(* IEC 61131-3 sources: plcc/demo/st-programs, 7 files *)

(* ---- alarm_system.st ---- *)
FUNCTION PriorityEncode : INT
VAR_INPUT critical : INT; high : INT; medium : INT; low : INT; END_VAR
    IF critical <> 0 THEN PriorityEncode := 4;
    ELSIF high <> 0 THEN PriorityEncode := 3;
    ELSIF medium <> 0 THEN PriorityEncode := 2;
    ELSIF low <> 0 THEN PriorityEncode := 1;
    ELSE PriorityEncode := 0;
    END_IF;
END_FUNCTION

FUNCTION_BLOCK AlarmHandler
VAR_INPUT
    temp_alarm : BOOL;
    pressure_alarm : BOOL;
    level_alarm : BOOL;
END_VAR
VAR_OUTPUT
    alarm_active : BOOL;
    alarm_code : INT;
END_VAR
VAR
    temp_val : INT;
    press_val : INT;
    level_val : INT;
END_VAR
    IF temp_alarm THEN temp_val := 1; ELSE temp_val := 0; END_IF;
    IF pressure_alarm THEN press_val := 1; ELSE press_val := 0; END_IF;
    IF level_alarm THEN level_val := 1; ELSE level_val := 0; END_IF;
    alarm_code := PriorityEncode(press_val, temp_val, level_val, 0);
    alarm_active := alarm_code > 0;
END_FUNCTION_BLOCK

PROGRAM AlarmSystem
VAR
    handler : AlarmHandler;
    system_alarm : BOOL;
    system_code : INT;
END_VAR
    handler(temp_alarm := TRUE, pressure_alarm := FALSE, level_alarm := TRUE);
    system_alarm := handler.alarm_active;
    system_code := handler.alarm_code;
END_PROGRAM

(* ---- motor_control.st ---- *)
FUNCTION_BLOCK MotorController
VAR_INPUT
    start_cmd : BOOL;
    stop_cmd : BOOL;
    current : REAL;
    overload_limit : REAL := 15.0;
END_VAR
VAR_OUTPUT
    running : BOOL;
    fault : BOOL;
    run_time : INT;
END_VAR
VAR
    overload_count : INT := 0;
END_VAR
    IF stop_cmd OR fault THEN
        running := FALSE;
    ELSIF start_cmd AND NOT fault THEN
        running := TRUE;
    END_IF;

    IF running THEN
        run_time := run_time + 1;
        IF current > overload_limit THEN
            overload_count := overload_count + 1;
            IF overload_count >= 3 THEN
                fault := TRUE;
                running := FALSE;
            END_IF;
        ELSE
            overload_count := 0;
        END_IF;
    END_IF;
END_FUNCTION_BLOCK

PROGRAM MotorSystem
VAR
    motor1 : MotorController;
    motor2 : MotorController;
    any_fault : BOOL;
END_VAR
    motor1(start_cmd := TRUE, stop_cmd := FALSE, current := 10.0);
    motor2(start_cmd := TRUE, stop_cmd := FALSE, current := 10.0);
    any_fault := motor1.fault OR motor2.fault;
END_PROGRAM

(* ---- pid_simple.st ---- *)
FUNCTION_BLOCK PID
VAR_INPUT
    setpoint : REAL;
    measured : REAL;
    kp : REAL := 1.0;
    ki : REAL := 0.1;
    kd : REAL := 0.05;
    dt : REAL := 0.01;
    out_min : REAL := -100.0;
    out_max : REAL := 100.0;
END_VAR
VAR_OUTPUT
    output : REAL;
END_VAR
VAR
    err : REAL;
    prev_err : REAL := 0.0;
    integral : REAL := 0.0;
    derivative : REAL;
END_VAR
    err := setpoint - measured;
    integral := integral + err * dt;
    derivative := (err - prev_err) / dt;
    output := kp * err + ki * integral + kd * derivative;

    (* Clamp output *)
    IF output > out_max THEN
        output := out_max;
    ELSIF output < out_min THEN
        output := out_min;
    END_IF;

    prev_err := err;
END_FUNCTION_BLOCK

PROGRAM PIDController
VAR
    pid_inst : PID;
    sensor_value : REAL := 0.0;
    target_value : REAL := 50.0;
    control_output : REAL;
END_VAR
    pid_inst(setpoint := target_value, measured := sensor_value);
    control_output := pid_inst.output;
END_PROGRAM

(* ---- water_treatment.st ---- *)
(* ═══════════════════════════════════════════════════════════ *)
(*  Water Treatment Plant — Industrial PLC Program            *)
(*  Registers 0-39 are SCADA-accessible via Modbus            *)
(* ═══════════════════════════════════════════════════════════ *)

(* ── Function Blocks ── *)

FUNCTION_BLOCK TankLevel
VAR_INPUT
    inlet_flow : REAL;
    outlet_flow : REAL;
    max_capacity : REAL;
END_VAR
VAR_OUTPUT
    level : REAL;
    level_pct : INT;
    high_alarm : BOOL;
    low_alarm : BOOL;
END_VAR
VAR
    high_sp : REAL := 90.0;
    low_sp : REAL := 10.0;
END_VAR
    level := level + (inlet_flow - outlet_flow) * 0.001;
    IF level < 0.0 THEN level := 0.0; END_IF;
    IF level > max_capacity THEN level := max_capacity; END_IF;
    level_pct := REAL_TO_INT(level * 100.0 / max_capacity);
    high_alarm := level_pct > 90;
    low_alarm := level_pct < 10;
END_FUNCTION_BLOCK

FUNCTION_BLOCK PumpControl
VAR_INPUT
    cmd_start : BOOL;
    cmd_stop : BOOL;
    speed_sp : INT;
    fault_reset : BOOL;
END_VAR
VAR_OUTPUT
    running : BOOL;
    speed : INT;
    fault : BOOL;
    hours : INT;
END_VAR
VAR
    scans : INT := 0;
END_VAR
    IF fault_reset THEN fault := FALSE; END_IF;
    IF cmd_stop THEN running := FALSE; END_IF;
    IF cmd_start AND NOT fault THEN running := TRUE; END_IF;
    IF running THEN
        speed := speed_sp;
        scans := scans + 1;
        hours := scans / 3600;
    ELSE
        speed := 0;
    END_IF;
END_FUNCTION_BLOCK

FUNCTION_BLOCK ValveControl
VAR_INPUT
    cmd_open : BOOL;
    cmd_close : BOOL;
END_VAR
VAR_OUTPUT
    position : INT;
    opened : BOOL;
    closed : BOOL;
END_VAR
    IF cmd_open AND NOT cmd_close THEN
        IF position < 100 THEN position := position + 5; END_IF;
    ELSIF cmd_close AND NOT cmd_open THEN
        IF position > 0 THEN position := position - 5; END_IF;
    END_IF;
    opened := position >= 100;
    closed := position <= 0;
END_FUNCTION_BLOCK

(* ── Main Program ── *)

PROGRAM WaterTreatment
VAR
    (* ═══════════════════════════════════════════ *)
    (* COMMANDS — write from SCADA (R0-R9)        *)
    (* ═══════════════════════════════════════════ *)
    cmd_start : INT := 0;         (* R0  write 1 to start *)
    cmd_stop : INT := 0;          (* R1  write 1 to stop *)
    cmd_flush : INT := 0;         (* R2  write 1 to flush *)
    cmd_alarm_ack : INT := 0;     (* R3  write 1 to acknowledge alarms *)
    cmd_alarm_reset : INT := 0;   (* R4  write 1 to reset faults *)
    sp_raw_tank : INT := 50;      (* R5  raw tank level setpoint % *)
    sp_clean_tank : INT := 70;    (* R6  clean tank level setpoint % *)
    sp_inlet_pump : INT := 60;    (* R7  inlet pump speed % *)
    sp_transfer_pump : INT := 40; (* R8  transfer pump speed % *)
    sp_outlet_pump : INT := 30;   (* R9  outlet pump speed % *)

    (* ═══════════════════════════════════════════ *)
    (* STATUS — read from SCADA (R10-R19)         *)
    (* ═══════════════════════════════════════════ *)
    running : INT := 0;           (* R10 process running *)
    stopped : INT := 1;           (* R11 process stopped *)
    flushing : INT := 0;          (* R12 flush in progress *)
    faulted : INT := 0;           (* R13 fault/alarm state *)
    cycle_count : INT := 0;       (* R14 scan counter *)
    raw_level : INT := 0;         (* R15 raw tank level % *)
    clean_level : INT := 0;       (* R16 clean tank level % *)
    system_ok : INT := 1;         (* R17 all systems healthy *)
    alarm_word : INT := 0;        (* R18 alarm bitmask *)
    total_flow : INT := 0;        (* R19 cumulative output *)

    (* ═══════════════════════════════════════════ *)
    (* EQUIPMENT STATUS (R20-R31)                 *)
    (* ═══════════════════════════════════════════ *)
    inlet_pump_run : INT := 0;    (* R20 *)
    inlet_pump_speed : INT := 0;  (* R21 *)
    inlet_pump_fault : INT := 0;  (* R22 *)
    xfer_pump_run : INT := 0;     (* R23 *)
    xfer_pump_speed : INT := 0;   (* R24 *)
    xfer_pump_fault : INT := 0;   (* R25 *)
    outlet_pump_run : INT := 0;   (* R26 *)
    outlet_pump_speed : INT := 0; (* R27 *)
    outlet_pump_fault : INT := 0; (* R28 *)
    inlet_vlv_pos : INT := 0;     (* R29 *)
    outlet_vlv_pos : INT := 0;    (* R30 *)
    drain_vlv_pos : INT := 0;     (* R31 *)

    (* ═══════════════════════════════════════════ *)
    (* ALARMS (R32-R39)                           *)
    (* ═══════════════════════════════════════════ *)
    alm_raw_high : INT := 0;      (* R32 raw tank high level *)
    alm_raw_low : INT := 0;       (* R33 raw tank low level *)
    alm_clean_high : INT := 0;    (* R34 clean tank high level *)
    alm_clean_low : INT := 0;     (* R35 clean tank low level *)
    alm_inlet_fault : INT := 0;   (* R36 inlet pump fault *)
    alm_xfer_fault : INT := 0;    (* R37 transfer pump fault *)
    alm_outlet_fault : INT := 0;  (* R38 outlet pump fault *)
    alm_count : INT := 0;         (* R39 total active alarms *)

    (* ═══════════════════════════════════════════ *)
    (* INTERNAL — FB instances after registers     *)
    (* ═══════════════════════════════════════════ *)
    raw_tank : TankLevel;
    clean_tank : TankLevel;
    p_inlet : PumpControl;
    p_transfer : PumpControl;
    p_outlet : PumpControl;
    v_inlet : ValveControl;
    v_outlet : ValveControl;
    v_drain : ValveControl;

    prev_running : INT := -1;
    init_done : INT := 0;
END_VAR

    (* ── Startup ── *)
    IF init_done = 0 THEN
        PRINT('Water Treatment PLC started');
        init_done := 1;
    END_IF;
    cycle_count := cycle_count + 1;

    (* ── Process commands (edge-triggered, auto-clear) ── *)
    IF cmd_start = 1 THEN
        cmd_start := 0;
        IF faulted = 0 THEN
            running := 1; stopped := 0; flushing := 0;
            PRINT('CMD: Process START');
        END_IF;
    END_IF;

    IF cmd_stop = 1 THEN
        cmd_stop := 0;
        running := 0; stopped := 1; flushing := 0;
        PRINT('CMD: Process STOP');
    END_IF;

    IF cmd_flush = 1 THEN
        cmd_flush := 0;
        running := 0; stopped := 0; flushing := 1;
        PRINT('CMD: FLUSH started');
    END_IF;

    IF cmd_alarm_ack = 1 THEN
        cmd_alarm_ack := 0;
        PRINT('CMD: Alarms acknowledged');
    END_IF;

    IF cmd_alarm_reset = 1 THEN
        cmd_alarm_reset := 0;
        faulted := 0;
        system_ok := 1;
        p_inlet(cmd_start := FALSE, cmd_stop := FALSE, speed_sp := 0, fault_reset := TRUE);
        p_transfer(cmd_start := FALSE, cmd_stop := FALSE, speed_sp := 0, fault_reset := TRUE);
        p_outlet(cmd_start := FALSE, cmd_stop := FALSE, speed_sp := 0, fault_reset := TRUE);
        PRINT('CMD: Faults reset');
    END_IF;

    (* ── Process control ── *)
    IF running = 1 THEN
        (* Inlet: fill raw tank to setpoint *)
        IF raw_level < sp_raw_tank THEN
            p_inlet(cmd_start := TRUE, cmd_stop := FALSE, speed_sp := sp_inlet_pump, fault_reset := FALSE);
            v_inlet(cmd_open := TRUE, cmd_close := FALSE);
        ELSE
            p_inlet(cmd_start := FALSE, cmd_stop := TRUE, speed_sp := 0, fault_reset := FALSE);
            v_inlet(cmd_open := FALSE, cmd_close := TRUE);
        END_IF;

        (* Transfer: move water from raw to clean *)
        IF raw_level > 20 AND clean_level < sp_clean_tank THEN
            p_transfer(cmd_start := TRUE, cmd_stop := FALSE, speed_sp := sp_transfer_pump, fault_reset := FALSE);
        ELSE
            p_transfer(cmd_start := FALSE, cmd_stop := TRUE, speed_sp := 0, fault_reset := FALSE);
        END_IF;

        (* Outlet: distribute clean water *)
        IF clean_level > 30 THEN
            p_outlet(cmd_start := TRUE, cmd_stop := FALSE, speed_sp := sp_outlet_pump, fault_reset := FALSE);
            v_outlet(cmd_open := TRUE, cmd_close := FALSE);
        ELSE
            p_outlet(cmd_start := FALSE, cmd_stop := TRUE, speed_sp := 0, fault_reset := FALSE);
            v_outlet(cmd_open := FALSE, cmd_close := TRUE);
        END_IF;

        v_drain(cmd_open := FALSE, cmd_close := TRUE);

    ELSIF flushing = 1 THEN
        (* Flush: drain everything *)
        p_inlet(cmd_start := FALSE, cmd_stop := TRUE, speed_sp := 0, fault_reset := FALSE);
        p_transfer(cmd_start := FALSE, cmd_stop := TRUE, speed_sp := 0, fault_reset := FALSE);
        p_outlet(cmd_start := FALSE, cmd_stop := TRUE, speed_sp := 0, fault_reset := FALSE);
        v_inlet(cmd_open := FALSE, cmd_close := TRUE);
        v_outlet(cmd_open := FALSE, cmd_close := TRUE);
        v_drain(cmd_open := TRUE, cmd_close := FALSE);

        (* Auto-stop flush when tanks are empty *)
        IF raw_level = 0 AND clean_level = 0 THEN
            flushing := 0; stopped := 1;
            PRINT('Flush complete');
        END_IF;

    ELSE
        (* Stopped / faulted *)
        p_inlet(cmd_start := FALSE, cmd_stop := TRUE, speed_sp := 0, fault_reset := FALSE);
        p_transfer(cmd_start := FALSE, cmd_stop := TRUE, speed_sp := 0, fault_reset := FALSE);
        p_outlet(cmd_start := FALSE, cmd_stop := TRUE, speed_sp := 0, fault_reset := FALSE);
        v_inlet(cmd_open := FALSE, cmd_close := TRUE);
        v_outlet(cmd_open := FALSE, cmd_close := TRUE);
        v_drain(cmd_open := FALSE, cmd_close := TRUE);
    END_IF;

    (* ── Tank simulation ── *)
    (* Flow rates scaled for demo speed — tanks fill in ~30 seconds *)
    raw_tank(
        inlet_flow := INT_TO_REAL(p_inlet.speed) * 50.0,
        outlet_flow := INT_TO_REAL(p_transfer.speed) * 30.0,
        max_capacity := 1000.0
    );
    clean_tank(
        inlet_flow := INT_TO_REAL(p_transfer.speed) * 30.0,
        outlet_flow := INT_TO_REAL(p_outlet.speed) * 20.0,
        max_capacity := 500.0
    );

    (* ── Copy to SCADA registers ── *)
    raw_level := raw_tank.level_pct;
    clean_level := clean_tank.level_pct;

    inlet_pump_run := BOOL_TO_INT(p_inlet.running);
    inlet_pump_speed := p_inlet.speed;
    inlet_pump_fault := BOOL_TO_INT(p_inlet.fault);

    xfer_pump_run := BOOL_TO_INT(p_transfer.running);
    xfer_pump_speed := p_transfer.speed;
    xfer_pump_fault := BOOL_TO_INT(p_transfer.fault);

    outlet_pump_run := BOOL_TO_INT(p_outlet.running);
    outlet_pump_speed := p_outlet.speed;
    outlet_pump_fault := BOOL_TO_INT(p_outlet.fault);

    inlet_vlv_pos := v_inlet.position;
    outlet_vlv_pos := v_outlet.position;
    drain_vlv_pos := v_drain.position;

    total_flow := total_flow + p_outlet.speed;

    (* ── Alarms ── *)
    alm_raw_high := BOOL_TO_INT(raw_tank.high_alarm);
    alm_raw_low := BOOL_TO_INT(raw_tank.low_alarm);
    alm_clean_high := BOOL_TO_INT(clean_tank.high_alarm);
    alm_clean_low := BOOL_TO_INT(clean_tank.low_alarm);
    alm_inlet_fault := BOOL_TO_INT(p_inlet.fault);
    alm_xfer_fault := BOOL_TO_INT(p_transfer.fault);
    alm_outlet_fault := BOOL_TO_INT(p_outlet.fault);

    (* Alarm word: bitmask of all active alarms *)
    alarm_word := alm_raw_high + alm_raw_low * 2 + alm_clean_high * 4
                + alm_clean_low * 8 + alm_inlet_fault * 16
                + alm_xfer_fault * 32 + alm_outlet_fault * 64;

    alm_count := alm_raw_high + alm_raw_low + alm_clean_high + alm_clean_low
               + alm_inlet_fault + alm_xfer_fault + alm_outlet_fault;

    (* Trip to fault only on critical alarms: high level or pump faults *)
    (* Low level alarms are informational — not a fault condition *)
    IF running = 1 THEN
        IF alm_raw_high = 1 OR alm_clean_high = 1 OR alm_inlet_fault = 1 OR alm_xfer_fault = 1 OR alm_outlet_fault = 1 THEN
            faulted := 1;
            running := 0;
            system_ok := 0;
            PRINT('FAULT: critical alarm, process stopped');
        END_IF;
    END_IF;

END_PROGRAM

(* ---- batch_process.st ---- *)
PROGRAM BatchProcess
VAR
    stage : INT := 0;
    timer : INT := 0;
    fill_valve : BOOL := FALSE;
    mixer : BOOL := FALSE;
    drain_valve : BOOL := FALSE;
    batch_count : INT := 0;
    complete : BOOL := FALSE;
END_VAR
    timer := timer + 1;
    CASE stage OF
        0: (* IDLE *)
            fill_valve := FALSE; mixer := FALSE; drain_valve := FALSE;
            stage := 1; timer := 0;
        1: (* FILL *)
            fill_valve := TRUE;
            IF timer >= 20 THEN stage := 2; timer := 0; fill_valve := FALSE; END_IF;
        2: (* MIX *)
            mixer := TRUE;
            IF timer >= 30 THEN stage := 3; timer := 0; mixer := FALSE; END_IF;
        3: (* DRAIN *)
            drain_valve := TRUE;
            IF timer >= 15 THEN
                stage := 0; timer := 0; drain_valve := FALSE;
                batch_count := batch_count + 1;
                complete := TRUE;
            END_IF;
    ELSE
        stage := 0;
    END_CASE;
END_PROGRAM

(* ---- blink.st ---- *)
PROGRAM Blink
VAR
    output : BOOL := FALSE;
END_VAR
    output := NOT output;
END_PROGRAM

(* ---- state_machine.st ---- *)
PROGRAM StateMachine
VAR
    state : INT := 0;
    output_a : BOOL := FALSE;
    output_b : BOOL := FALSE;
    input_trigger : BOOL := FALSE;
    counter : INT := 0;
END_VAR
    CASE state OF
        0:
            output_a := FALSE;
            output_b := FALSE;
            IF input_trigger THEN
                state := 1;
            END_IF;
        1:
            output_a := TRUE;
            output_b := FALSE;
            counter := counter + 1;
            IF counter >= 10 THEN
                state := 2;
                counter := 0;
            END_IF;
        2:
            output_a := FALSE;
            output_b := TRUE;
            counter := counter + 1;
            IF counter >= 5 THEN
                state := 0;
                counter := 0;
            END_IF;
    ELSE
        state := 0;
    END_CASE;
END_PROGRAM
